FUNCTION FC 1 : VOID
BEGIN
NETWORK
TITLE Lamp
END_FUNCTION
